Fanuc KAREL source: KT00832.KL

PROGRAM KT00832
%NOLOCKGROUP
VAR
  I1: INTEGER
  I2: INTEGER
  OUT: INTEGER
BEGIN
  I1 = 2
  I2 = 3
  I1 = 2
  I2 = 3
  OUT = SQRT(I1)
END KT00832
